ABB RobotStudio station: 项目2.rsstn

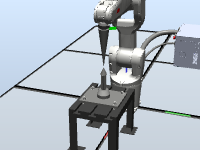
Station Station (saved by RobotStudio 6.8.8148.134)
Controller test2
  mechanical unit ROB_1: IRB1200_5_90_STD_02, 6 joints, base frame (0, 0, 0) mm
Layout (positions relative to the parent item):
  - IRB1200_5_90_STD_02 [mechanism, from Robots\IRB1200_5_90_STD_02.rslib] at (0, 0, 0) mm; joint values [0.0005, 0.145, -0.0543, -0.001, 1.4815, -0.576] (rad or m)
  - table_and_fixture_140 [part, from Training Objects\propeller_table.rslib] at (292.73, -175, 0) mm
  - IRC5_Compact [part, from Equipment\IRC5_Compact__02.rslib] at (-1366.51, 213.23, 0) mm
  - PhysicsCable_1 [physicscable]
  - PhysicsCable_2 [physicscable]
  - 部件_1 [part]
  - 部件_2 [part] at (517.58, 0.15, 761.34) mm, rotated rx -180 ry -0.11 rz -146.96 deg
Attachment: 部件_2 is attached to IRB1200_5_90_STD_02 / Link6
Targets, tools, work objects and paths stored in the station, written as RAPID:
! task T_ROB1
MODULE Module1
  PERS tooldata tool1:=[TRUE,[[0,0,0],[1,0,0,0]],[1,[0,0,10],[1,0,0,0],0,0,0]];
ENDMODULE

